Fanuc KAREL source: kd00068.KL

-- PROVISIONAL review KL for V940-1; original PC SHA256 185527df14943be4de279c40240d03046571e8006072339d1a577fa61ab104a2
-- Incomplete behavior may be omitted. Consult companion uncertainty JSON. Do not deploy.
PROGRAM KD00068
%NOLOCKGROUP
VAR
  I : INTEGER
  J : INTEGER
  B : BOOLEAN
  R : REAL
  S : STRING[80]
BEGIN
  -- V9_ZERO_TABLE_METADATA_HINT layout=0001; no indexed target words; source/name/runtime held
  -- UNRESOLVED_PC offsets 5-29; opcodes 9D,81,18,9D,1B,9D,12,2E,1B,2E,13,04
  -- UNRESOLVED_PC offsets 34-38; opcodes 7F
END KD00068
